FUNCTION_BLOCK Testing_HMI (* Service Interface Function Block Type *)
  (* Standard: 61499-2 *)
  (* Version 0.0, 11/16/2026, Sandeep Patil, Flexbridge AB, template *)
  PACKAGE Flexbridge.FestoMPS400;
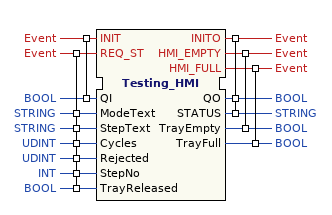
  EVENT_INPUT
    INIT WITH QI;
    REQ_ST WITH ModeText, StepText, Cycles, Rejected, StepNo, TrayReleased;
  END_EVENT
  EVENT_OUTPUT
    INITO WITH QO, STATUS;
    HMI_EMPTY WITH TrayEmpty;
    HMI_FULL WITH TrayFull;
  END_EVENT
  VAR_INPUT
    QI : BOOL; (* Input event qualifier *)
    ModeText : STRING; (* Station mode *)
    StepText : STRING; (* Current step (number and name) *)
    Cycles : UDINT; (* Workpieces put on a tray since start-up *)
    Rejected : UDINT; (* Workpieces rejected since start-up *)
    StepNo : INT; (* Current step number *)
    TrayReleased : BOOL; (* The tray has been released (until the next tray) *)
  END_VAR
  VAR_OUTPUT
    QO : BOOL; (* Event Output Qualifier *)
    STATUS : STRING; (* Service Status *)
    TrayEmpty : BOOL; (* Stand-in button: an empty tray has arrived at interface 1 *)
    TrayFull : BOOL; (* Stand-in button: a tray with a workpiece has arrived at interface 1 *)
  END_VAR
  SERVICE /
    SEQUENCE 
    END_SEQUENCE
  END_SERVICE
END_FUNCTION_BLOCK
